// TIA Portal V21 export
TextList "TL_Phase"  ListRange=Decimal
  TextListEntry   Text="vožnja do izvora"
  TextListEntry   From=1, To=1, Text="podizanje"
  TextListEntry   From=2, To=2, Text="vožnja do odredišta"
  TextListEntry   From=3, To=3, Text="spuštanje"
